(* IEC 61131-3 sources: IRIS-Project/LASAL CONTROL SOFTWARE/LasalProject_2025_09_12/Network/Timer, 1 file *)

(* ---- ONE_Timer_Table.st ---- *)
#define OBJECTS_CONFIG

FUNCTION GLOBAL TAB ONE_Timer
-1$UINT, 0$UINT,
0$UINT, 0$UINT,

7$UDINT,
TO_UDINT(1642197576), "DischargeTimer", 0$UINT, 0$UINT, 1$UINT,
TO_UDINT(2171929650), "IrradiationManager", 0$UINT, 0$UINT, 1$UINT,
TO_UDINT(2103413850), "MoveTimer", 0$UINT, 0$UINT, 1$UINT,
TO_UDINT(2815000061), "Reset", 0$UINT, 0$UINT, 1$UINT,
TO_UDINT(3035062039), "SysDateTime", 1$UINT, 5$UINT, 3$UINT,
TO_UDINT(1512043018), "TimeDateLib", 1$UINT, 1$UINT, 3$UINT,
TO_UDINT(3890592521), "TimerLib", 1$UINT, 0$UINT, 3$UINT,

_NO_ATTR, TO_UDINT(4223322087), "DISCHARGETIMER1",

_NO_ATTR, TO_UDINT(101499717), "IRRADIATIONTIMERS",

_NO_ATTR, TO_UDINT(136251601), "MOVETIMER1",

_NO_ATTR, TO_UDINT(1081583723), "RESET1",

_NO_ATTR, TO_UDINT(12291375), "SYSDATETIME1",
_NO_ATTR, TO_UDINT(2578635925), "SYSDATETIME2",
_NO_ATTR, TO_UDINT(4004899843), "SYSDATETIME3",

_NO_ATTR, TO_UDINT(1666390363), "TIMEDATELIB1",
_NO_ATTR, TO_UDINT(1693608047), "TIMEDATELIB1_COPY",
_NO_ATTR, TO_UDINT(4200220897), "TIMEDATELIB2",

_NO_ATTR, TO_UDINT(4209488552), "TIMERLIB1",
_NO_ATTR, TO_UDINT(2480454521), "TIMERLIB1_COPY",
_NO_ATTR, TO_UDINT(3243102297), "TIMERLIB1_COPY_COPY",

//Internal connections
0$UDINT,
0$UDINT,
0$UDINT,
14$UDINT,
TO_UDINT(0), "c_timer", TO_UDINT(7), "ClassSvr",
TO_UDINT(0), "c_SysDate", TO_UDINT(4), "SysDate",
TO_UDINT(0), "c_SysTime", TO_UDINT(4), "SysTime",
TO_UDINT(1), "Timer1", TO_UDINT(10), "ClassSvr",
TO_UDINT(1), "Timer2", TO_UDINT(11), "ClassSvr",
TO_UDINT(1), "Timer3", TO_UDINT(12), "ClassSvr",
TO_UDINT(1), "c_timerLib", TO_UDINT(8), "ClassSvr",
TO_UDINT(1), "c_SysTime", TO_UDINT(6), "SysTime",
TO_UDINT(2), "c_timer", TO_UDINT(9), "ClassSvr",
TO_UDINT(2), "c_SysDate", TO_UDINT(5), "SysDate",
TO_UDINT(2), "c_SysTime", TO_UDINT(5), "SysTime",
TO_UDINT(3), "c_ResetTimerIrr", TO_UDINT(1), "s_Reset",
TO_UDINT(3), "c_ResetTimerMov", TO_UDINT(2), "s_Reset",
TO_UDINT(3), "c_ResetTimerDis", TO_UDINT(0), "s_Reset",

//Initialization values
0$UDINT,
1$UDINT,
TO_UDINT(0), "c_timer", TO_UDINT(0),//|Timer.DischargeTimer1.c_timer;

//Symbolic initialization values
0$UDINT,
0$UDINT,

//Initialization of string values
0$UDINT,
0$UDINT,

//Configuration of tasks (RealTime, Cyclic, Background)
0$UDINT,
0$UDINT,

0$UDINT,
7$UDINT,
TO_UDINT(0), (100)$UDINT, 4194303$DINT, 	//DISCHARGETIMER1
TO_UDINT(1), (100)$UDINT, 4194303$DINT, 	//IRRADIATIONTIMERS
TO_UDINT(2), (100)$UDINT, 4194303$DINT, 	//MOVETIMER1
TO_UDINT(3), (100)$UDINT, 4194303$DINT, 	//RESET1
TO_UDINT(4), (-2147483148)$UDINT, 4194303$DINT, 	//SYSDATETIME1
TO_UDINT(5), (-2147483148)$UDINT, 4194303$DINT, 	//SYSDATETIME2
TO_UDINT(6), (-2147483148)$UDINT, 4194303$DINT, 	//SYSDATETIME3

0$UDINT,
0$UDINT,

//External connections
0$UDINT,
3$UDINT,
TO_UDINT(1), "TabletInIrrPos", C_DIR, TO_UDINT(593259826), "Motore_M51","s_tablet_irradiation_position",
TO_UDINT(1), "NrIrrTablets", C_DIR, TO_UDINT(593259826), "Motore_M51","s_TabletTimer",
TO_UDINT(1), "SetStartStopIrr", C_DIR, TO_UDINT(1533940179), "Manager_globale1","ComandoIrradiation",

//Magic internal connections
0$UDINT,
0$UDINT,

//Configuration of timeslots of tasks (RealTime, Cyclic)
#ifdef __LSLLDR_TIMESLOTS__
0$UDINT,
0$UDINT,

0$UDINT,
0$UDINT,

#endif //__LSLLDR_TIMESLOTS__

//MultiMaster connections
#ifdef __LSLLDR_MULTIMASTER__
0$UDINT,
0$UDINT,
#endif //__LSLLDR_MULTIMASTER__

//Configuration for task ID (RealTime, CyclicTime)
#ifdef __LSLLDR_TASKID__
"\\\\TASKS2  "
0$UDINT,
0$UDINT,

0$UDINT,
7$UDINT,
(0)$UDINT, 	//DISCHARGETIMER1
(0)$UDINT, 	//IRRADIATIONTIMERS
(0)$UDINT, 	//MOVETIMER1
(0)$UDINT, 	//RESET1
(0)$UDINT, 	//SYSDATETIME1
(0)$UDINT, 	//SYSDATETIME2
(0)$UDINT, 	//SYSDATETIME3

0$UDINT,
0$UDINT,

#endif //__LSLLDR_TASKID__

END_FUNCTION
